(* IEC 61131-3 sources: kns-port-domestic/upstream/kns-pump-station/src/POUs/Model/FB_HydraulicSolver, 6 files *)

(* ---- FB_HydraulicSolver.decl.st ---- *)
// Назначение: рабочая точка насосов на общий напорный коллектор по законам подобия. Насос:
//             H_i = H0·s_i² − k_i·q_i², s = f / 50 Гц; сеть: H = (Hgeo − h) + R·Q², Q = Σ q_i; обратные
//             клапаны — q_i = 0 при H0·s_i² ≤ H. Напор — бисекцией на [Hgeo − h, max(H0·s_i²)]
//             (SIM_SOLVER_ITERATIONS шагов): так решаются и разные частоты. Сухой ход насоса и
//             осушенный приёмок — подача 0 и ток холостого хода; засор — k_i·SIM_CLOG_K_FACTOR, ток
//             ×SIM_CLOG_I_FACTOR к току того же насоса в сети без засора (второе решение; только у насоса,
//             который может подавать). Давление PT201 (у дна, условно):
//             ρ·g·(H + h)/10⁵ бар; насосы стоят — столб за обратными клапанами ρ·g·Hgeo/10⁵.
// Автор:      kr0nsch
// Версия:     0.1.1
// Документ:   docs/DESIGN.md, разделы 11.2, 11.3; эталон tools_project/plant_reference.py
FUNCTION_BLOCK FB_HydraulicSolver
VAR_INPUT
    arSpeed    : ARRAY[1..GVL_Const.STN_PUMP_COUNT] OF REAL;   // s = f / 50 Гц; ≤ 0 — насос не вращается
    axAirLock  : ARRAY[1..GVL_Const.STN_PUMP_COUNT] OF BOOL;   // сухой ход насоса (stFaultInj.axAirLock)
    axClog     : ARRAY[1..GVL_Const.STN_PUMP_COUNT] OF BOOL;   // засор (stFaultInj.axClog)
    rLevel_m   : REAL;              // уровень в резервуаре
    xIntakeDry : BOOL;              // приёмок осушен (FB_TankModel.xIntakeDry)
    stPump     : ST_PumpModelCfg;   // характеристика насоса и сети
END_VAR
VAR_OUTPUT
    arFlow_m3h   : ARRAY[1..GVL_Const.STN_PUMP_COUNT] OF REAL;   // подачи насосов
    arCurrent_A  : ARRAY[1..GVL_Const.STN_PUMP_COUNT] OF REAL;   // токи двигателей
    rFlow_m3h    : REAL;            // подача станции (FT202)
    rHead_m      : REAL;            // напор сети
    rPressure_bar : REAL;           // давление в коллекторе (PT201)
END_VAR
VAR
    arQ        : ARRAY[1..GVL_Const.STN_PUMP_COUNT] OF REAL;   // подачи последнего решения Solve
    arShutoff  : ARRAY[1..GVL_Const.STN_PUMP_COUNT] OF REAL;   // H0·s² (напор при закрытой задвижке)
    arK        : ARRAY[1..GVL_Const.STN_PUMP_COUNT] OF REAL;   // действующая крутизна
    axActive   : ARRAY[1..GVL_Const.STN_PUMP_COUNT] OF BOOL;   // насос может подавать
    arS        : ARRAY[1..GVL_Const.STN_PUMP_COUNT] OF REAL;   // скорость после проверки
    xAnyClog   : BOOL;              // есть подающий насос с засором (нужно второе решение)
    rHeadClean : REAL;              // напор сети без засоров
    uiPump     : UINT;              // индекс насоса
END_VAR

(* ---- FB_HydraulicSolver.impl.st ---- *)
// 1. Скорости (неконечная — как 0) и какие насосы могут подавать
xAnyClog := FALSE;
FOR uiPump := 1 TO GVL_Const.STN_PUMP_COUNT DO
    IF PL.F_IsFinite(rIn := arSpeed[uiPump]) AND arSpeed[uiPump] > 0.0 THEN
        arS[uiPump] := arSpeed[uiPump];
    ELSE
        arS[uiPump] := 0.0;
    END_IF
    axActive[uiPump] := arS[uiPump] > 0.0 AND NOT axAirLock[uiPump] AND NOT xIntakeDry;
    arShutoff[uiPump] := stPump.rH0_m * arS[uiPump] * arS[uiPump];
    xAnyClog := xAnyClog OR (axClog[uiPump] AND axActive[uiPump]);
END_FOR

// 2. Рабочая точка с засорами и токи по ней
rHead_m := Solve(xWithClog := TRUE);
rFlow_m3h := 0.0;
FOR uiPump := 1 TO GVL_Const.STN_PUMP_COUNT DO
    arFlow_m3h[uiPump] := arQ[uiPump];
    rFlow_m3h := rFlow_m3h + arQ[uiPump];
    arCurrent_A[uiPump] := F_PumpCurrent(rFlow_m3h := arQ[uiPump], rHead_m := rHead_m, rSpeed := arS[uiPump],
                                         stPump := stPump);
END_FOR

// 3. Засор: ток ×SIM_CLOG_I_FACTOR к току того же насоса в той же сети без засора — только у насоса, который
//    может подавать (при сухом ходе и осушенном приёмке воды в колесе нет: ток холостого хода, ниже порога
//    недогрузки)
IF xAnyClog THEN
    rHeadClean := Solve(xWithClog := FALSE);
    FOR uiPump := 1 TO GVL_Const.STN_PUMP_COUNT DO
        IF axClog[uiPump] AND axActive[uiPump] THEN
            arCurrent_A[uiPump] := GVL_Const.SIM_CLOG_I_FACTOR
                                   * F_PumpCurrent(rFlow_m3h := arQ[uiPump], rHead_m := rHeadClean,
                                                   rSpeed := arS[uiPump], stPump := stPump);
        END_IF
    END_FOR
END_IF

// 4. Давление у дна коллектора: напор сети плюс уровень
rPressure_bar := GVL_Const.SIM_RHO_KGM3 * GVL_Const.SIM_GRAVITY_MPS2 * (rHead_m + rLevel_m) / GVL_Const.SIM_PA_PER_BAR;

(* ---- FlowsAt.method.decl.st ---- *)
// Подачи насосов при напоре rHead_m (в arQ): √((H0·s² − H)/k) для насосов, которые могут подавать
// и открывают обратный клапан; результат — сумма
METHOD PRIVATE FlowsAt : REAL
VAR_INPUT
    rHead_m : REAL;         // напор сети
END_VAR
VAR
    uiJ : UINT;             // индекс насоса
END_VAR

(* ---- FlowsAt.method.impl.st ---- *)
FlowsAt := 0.0;
FOR uiJ := 1 TO GVL_Const.STN_PUMP_COUNT DO
    IF axActive[uiJ] AND arShutoff[uiJ] > rHead_m AND arK[uiJ] > 0.0 THEN
        arQ[uiJ] := SQRT((arShutoff[uiJ] - rHead_m) / arK[uiJ]);
    ELSE
        arQ[uiJ] := 0.0;
    END_IF
    FlowsAt := FlowsAt + arQ[uiJ];
END_FOR

(* ---- Solve.method.decl.st ---- *)
// Напор сети в рабочей точке (бисекция по H); подачи — в arQ. xWithClog = FALSE — как будто
// засоров нет (для тока засорённого насоса). Нет насоса, способного преодолеть статический напор, —
// подачи 0, напор Hgeo − h
METHOD PRIVATE Solve : REAL
VAR_INPUT
    xWithClog : BOOL;       // учитывать засоры
END_VAR
VAR
    rStatic : REAL;         // статический напор Hgeo − h
    rLo     : REAL;         // границы бисекции по напору
    rHi     : REAL;
    rMid    : REAL;
    rTotal  : REAL;         // подача станции при rMid
    uiIter  : UINT;         // шаг бисекции
    uiI     : UINT;         // индекс насоса
END_VAR

(* ---- Solve.method.impl.st ---- *)
rStatic := stPump.rHgeo_m - rLevel_m;
rHi := rStatic;
FOR uiI := 1 TO GVL_Const.STN_PUMP_COUNT DO
    arQ[uiI] := 0.0;
    IF xWithClog AND axClog[uiI] THEN
        arK[uiI] := stPump.rK_mh2 * GVL_Const.SIM_CLOG_K_FACTOR;
    ELSE
        arK[uiI] := stPump.rK_mh2;
    END_IF
    IF axActive[uiI] AND arShutoff[uiI] > rHi THEN
        rHi := arShutoff[uiI];
    END_IF
END_FOR

// ни один насос не преодолевает статический напор (или характеристика неверна) — обратные клапаны закрыты
IF rHi <= rStatic OR stPump.rK_mh2 <= 0.0 OR stPump.rR_mh2 < 0.0 THEN
    Solve := rStatic;
    RETURN;
END_IF

// f(H) = Hst + R·Q(H)² − H убывает по H: f(Hst) ≥ 0, f(max H0·s²) < 0
rLo := rStatic;
FOR uiIter := 1 TO GVL_Const.SIM_SOLVER_ITERATIONS DO
    rMid := (rLo + rHi) / 2.0;
    rTotal := FlowsAt(rHead_m := rMid);
    IF rStatic + stPump.rR_mh2 * rTotal * rTotal > rMid THEN
        rLo := rMid;
    ELSE
        rHi := rMid;
    END_IF
END_FOR
Solve := (rLo + rHi) / 2.0;
rTotal := FlowsAt(rHead_m := Solve);
